(* IEC 61131-3 sources: 2026_Projet_YGO_ExcavatriceDragage/CODE_BACKUP/CODE_20260904_AvantWeekendBackup_v0.6.34/A_COMMUN/_TYPES, 6 files *)

(* ---- E_State.st ---- *)
(* =======================================================================
   ⚙️ E_State — Phase opérationnelle d'un FB métier (valeurs EXCLUSIVES)
   ───────────────────────────────────────────────────────────────
   🎯 Rôle : Énumération des phases opérationnelles d'un FB métier
   ⚙️ Machine d'état : Un seul état actif à la fois (orthogonal à Error)
   📄 Doc métier : DOC/AF/AF_Partie-03_Contrats_Composants_v2.3.md §3
   ======================================================================= *)

TYPE E_State :
ENUM
    DISABLED := 0,   (* Enable faux, neutralisé *)
    INIT     := 1,   (* Démarrage / vérifs *)
    READY    := 2,   (* Prêt, attend ordre *)
    BUSY     := 3,   (* Action en cours *)
    DONE     := 4,   (* Action terminée *)
    STOPPING := 5,   (* Décél rampe avant arrêt (StartStop=FALSE ou SafeStop=TRUE) *)
    ERROR    := 6    (* Défaut actif non acquitté (FB en erreur — HMI non aveugle) *)
END_ENUM
END_TYPE

(* ---- ST_ContactorCheck.st ---- *)
(* =======================================================================
   🔌 ST_ContactorCheck — Double vérification commande/retour contacteur
   ───────────────────────────────────────────────────────────────
   🎯 Rôle : Structure de diagnostic pour vérification commande vs retour
   📊 Diagnostic : Détection des défauts contacteur (StuckClosed / StuckOpen)
   📄 Doc métier : DOC/AF/AF_Partie-03_Contrats_Composants_v2.3.md §2
   ======================================================================= *)

TYPE ST_ContactorCheck :
STRUCT
    Command     : BOOL;   // Ordre envoyé au contacteur (TRUE = fermé/actif)
    Feedback    : BOOL;   // Retour d'état câblé (TRUE = effectivement fermé)
    StuckClosed : BOOL;   // Diag : commande OFF mais retour ON depuis trop longtemps → PowerCutOff
    StuckOpen   : BOOL;   // Diag : commande ON mais retour OFF depuis trop longtemps
END_STRUCT
END_TYPE

(* ---- ST_Fault.st ---- *)
(* =======================================================================
   🧩 ST_Fault — Brique socle défaut (2 vues : live + latchée)
   ───────────────────────────────────────────────────────────────
   🎯 Rôle : porter l'état défaut d'un composant, applicable dans TOUS les cas
      (acquittable ou non), sans brique warning séparée.
        • Vue LIVE   (Error / ErrorId)     : suit la cause, retombe seule à 0.
        • Vue LATCHÉE (Latched / LatchedId): mémorisée au défaut, reste jusqu'au front Reset.
      Le choix acquittable / non-acquittable se fait PAR CAUSE
      (ST_FaultCause.Latching), jamais par bloc.
   🔒 Sécurité : interlock TOUJOURS sur la cause brute (Error / ErrorId), jamais
      sur l'acquittement. Reset TOUJOURS effectif, jamais conditionné (std §9).
   🧬 Composition : brique de base réutilisable — sortie de FB, struct métier, GVL.
      Texte IHM NON stocké ici : dérivé côté IHM depuis LatchedId / ErrorId.
   📄 Doc : DOC/STDS/CODE_QUALITY_STANDARDS.md §2quinquies / §9
   ======================================================================= *)

TYPE ST_Fault :
STRUCT
    Error     : BOOL;   (* <-- [DIAG] vue LIVE : au moins une cause présente maintenant *)
    ErrorId   : WORD;    (* <-- [DIAG] bitfield des causes présentes maintenant (0 si aucune) *)
    Latched   : BOOL;    (* <-- [DIAG] vue LATCHÉE : défaut non acquitté, reste jusqu'au front Reset *)
    LatchedId : WORD;    (* <-- [DIAG] ErrorId figé à l'apparition du défaut, effacé au Reset *)
END_STRUCT
END_TYPE

(* ---- ST_FaultCause.st ---- *)
(* =======================================================================
   🧩 ST_FaultCause — Cause élémentaire alimentant ST_Fault (socle FB_FaultCore)
   ───────────────────────────────────────────────────────────────
   🎯 Rôle : une cause exprimée EN CLAIR (BOOL + libellé), sans bitfield ni masque.
      Le FB métier remplit une liste (ARRAY[0..15] OF ST_FaultCause) ;
      le socle FB_FaultCore en déduit ST_Fault (vue live + vue latchée).
   🔒 Sécurité : interlock TOUJOURS sur Active (cause brute), jamais sur le latch.
      Latching = TRUE  → la cause ARME la vue latchée (défaut à acquitter).
      Latching = FALSE → la cause n'alimente que la vue live (retombe seule).
      Fail-safe : une cause laissée à Latching=FALSE reste visible en live —
      pour la rendre acquittable, il faut le déclarer explicitement.
   📄 Doc : DOC/STDS/CODE_QUALITY_STANDARDS.md §2quinquies / §9
   ======================================================================= *)

TYPE ST_FaultCause :
STRUCT
    Active   : BOOL;    (* 1 = cause présente maintenant (interlock sur cette valeur) *)
    Latching : BOOL;    (* 1 = cause à acquitter (arme Latched) ; 0 = live seulement *)
    Texte    : STRING;  (* libellé prêt IHM (non stocké dans ST_Fault, dérivé côté IHM) *)
END_STRUCT
END_TYPE

(* ---- ST_Lifecycle.st ---- *)
(* =======================================================================
   🧩 ST_Lifecycle — Brique socle cycle d'exécution
   ───────────────────────────────────────────────────────────────
   🎯 Rôle : porter l'avancement d'une action à cycle (organe, séquenceur).
      Optionnelle : un FB purement synchrone (conditionneur, filtre, joystick)
      ne la porte pas.
   🧬 Composition : brique de base réutilisable, composée avec ST_Fault.
   📄 Doc : DOC/STDS/CODE_QUALITY_STANDARDS.md §2quinquies
   ======================================================================= *)

TYPE ST_Lifecycle :
STRUCT
    Busy : BOOL;   (* <-- [STAT] 1 = action en cours *)
    Done : BOOL;   (* <-- [STAT] 1 = action terminée avec succès *)
END_STRUCT
END_TYPE

(* ---- ST_Status.st ---- *)
(* =======================================================================
   🧩 ST_Status — Socle transverse de statut d'un FB métier
   ───────────────────────────────────────────────────────────────
   🎯 Rôle : regroupe l'état, le défaut et le warning d'un FB standard,
      avec les textes prêts pour l'IHM (plus de conditions complexes
      côté affichage). Évolution additive : les 6 membres d'origine sont conservés.
   🧬 Forme cible : les FB standard exposent `Status : ST_Status`
      rempli via le socle `FB_FbStatus` (même comportement partout).
   ⚠️ State/StateAtError : E_State (phases opérationnelles FB métier).
      Un FB dont l'état est un énum domaine (E_Diag_State, CycleStep,
      ST_Safety_Emergency_State…) garde sa sortie typée SÉPARÉE et ne
      migre pas vers ST_Status (exception documentée).
   📄 Doc : DOC/STDS/CODE_QUALITY_STANDARDS.md §2quinquies
   ======================================================================= *)

TYPE ST_Status :
STRUCT
    (* ---- membres historiques (conservés) ---- *)
    Busy         : BOOL;    (* 1 = Bloc en cours d'exécution *)
    Done         : BOOL;    (* 1 = Action terminée avec succès *)
    Error        : BOOL;    (* 1 = Défaut à acquitter (laté jusqu'au Reset) *)
    ErrorId      : WORD;    (* Code d'erreur bitfield / enum diagnostic *)
    State        : E_State; (* État courant de la machine d'état *)
    StateAtError : E_State; (* État mémorisé lors de l'apparition du défaut *)
    (* ---- membres ajoutés (forme cible enrichie) ---- *)
    Warning        : BOOL;  (* 1 = warning actif (auto-effacé, aucun acquittement) *)
    WarningId      : WORD;  (* Code warning courant (bitfield) *)
    WarningIdTxt   : STRING;(* Texte généré depuis WarningId (prêt IHM) *)
    ErrorIdTxt     : STRING;(* Texte généré depuis ErrorId *)
    ResetRequested : BOOL;  (* 1 = un Reset est nécessaire / en cours *)
END_STRUCT
END_TYPE
